(* PLC project GeneratedProgram, SafePLC-Gen SafePLC-Gen Multimodal 1.0 *)
(* stored: creationDateTime 2026-04-25T12:15:41.761626Z *)

PROGRAM GeneratedProgram
  VAR
    TI_2909_Scaled : REAL;
    TT_2909_Scaled : REAL;
    TT_2911_Scaled : REAL;
    TT_2917_Scaled : REAL;
    TI_2917_Scaled : REAL;
    XI_2901A_Scaled : REAL;
    XI_2901B_Scaled : REAL;
    TI_2909_HH_SP : REAL;
    TI_2909_H_SP : REAL;
    TI_2909_L_SP : REAL;
    TI_2909_LL_SP : REAL;
    TI_2909_Deadband : REAL;
    TI_2909_HH : BOOL;
    TI_2909_H : BOOL;
    TI_2909_L : BOOL;
    TI_2909_LL : BOOL;
    TI_2909_HH_Latch : SR;
    TI_2909_LL_Latch : SR;
    TI_2909_HH_Ack : BOOL;
    TI_2909_LL_Ack : BOOL;
    TT_2909_HH_SP : REAL;
    TT_2909_H_SP : REAL;
    TT_2909_L_SP : REAL;
    TT_2909_LL_SP : REAL;
    TT_2909_Deadband : REAL;
    TT_2909_HH : BOOL;
    TT_2909_H : BOOL;
    TT_2909_L : BOOL;
    TT_2909_LL : BOOL;
    TT_2909_HH_Latch : SR;
    TT_2909_LL_Latch : SR;
    TT_2909_HH_Ack : BOOL;
    TT_2909_LL_Ack : BOOL;
    TT_2911_HH_SP : REAL;
    TT_2911_H_SP : REAL;
    TT_2911_L_SP : REAL;
    TT_2911_LL_SP : REAL;
    TT_2911_Deadband : REAL;
    TT_2911_HH : BOOL;
    TT_2911_H : BOOL;
    TT_2911_L : BOOL;
    TT_2911_LL : BOOL;
    TT_2911_HH_Latch : SR;
    TT_2911_LL_Latch : SR;
    TT_2911_HH_Ack : BOOL;
    TT_2911_LL_Ack : BOOL;
    TIC_2911_SP : REAL;
    TIC_2911_Kp : REAL;
    TIC_2911_Ki : REAL;
    TIC_2911_Error : REAL;
    TIC_2911_Integral : REAL;
    TIC_2911_Output : REAL;
    TT_2917_HH_SP : REAL;
    TT_2917_H_SP : REAL;
    TT_2917_L_SP : REAL;
    TT_2917_LL_SP : REAL;
    TT_2917_Deadband : REAL;
    TT_2917_HH : BOOL;
    TT_2917_H : BOOL;
    TT_2917_L : BOOL;
    TT_2917_LL : BOOL;
    TT_2917_HH_Latch : SR;
    TT_2917_LL_Latch : SR;
    TT_2917_HH_Ack : BOOL;
    TT_2917_LL_Ack : BOOL;
    TI_2917_HH_SP : REAL;
    TI_2917_H_SP : REAL;
    TI_2917_L_SP : REAL;
    TI_2917_LL_SP : REAL;
    TI_2917_Deadband : REAL;
    TI_2917_HH : BOOL;
    TI_2917_H : BOOL;
    TI_2917_L : BOOL;
    TI_2917_LL : BOOL;
    TI_2917_HH_Latch : SR;
    TI_2917_LL_Latch : SR;
    TI_2917_HH_Ack : BOOL;
    TI_2917_LL_Ack : BOOL;
    XI_2901A_HH_SP : REAL;
    XI_2901A_H_SP : REAL;
    XI_2901A_L_SP : REAL;
    XI_2901A_LL_SP : REAL;
    XI_2901A_Deadband : REAL;
    XI_2901A_HH : BOOL;
    XI_2901A_H : BOOL;
    XI_2901A_L : BOOL;
    XI_2901A_LL : BOOL;
    XI_2901A_HH_Latch : SR;
    XI_2901A_LL_Latch : SR;
    XI_2901A_HH_Ack : BOOL;
    XI_2901A_LL_Ack : BOOL;
    XI_2901B_HH_SP : REAL;
    XI_2901B_H_SP : REAL;
    XI_2901B_L_SP : REAL;
    XI_2901B_LL_SP : REAL;
    XI_2901B_Deadband : REAL;
    XI_2901B_HH : BOOL;
    XI_2901B_H : BOOL;
    XI_2901B_L : BOOL;
    XI_2901B_LL : BOOL;
    XI_2901B_HH_Latch : SR;
    XI_2901B_LL_Latch : SR;
    XI_2901B_HH_Ack : BOOL;
    XI_2901B_LL_Ack : BOOL;
    LOOP_2917_TRIP : BOOL;
    LOOP_2901A_TRIP : BOOL;
    LOOP_2901B_TRIP : BOOL;
    LOOP_3200_TRIP : BOOL;
    TT_2917_HH_Trip : BOOL;
    TT_2917_LL_Trip : BOOL;
    VSHH_2901A_HH : BOOL;
    VSHH_2901A_LL : BOOL;
    VSHH_2901B_HH : BOOL;
    VSHH_2901B_LL : BOOL;
    ESD_3200_HH : BOOL;
    ESD_3200_LL : BOOL;
    SAFE_STATE : BOOL;
    MotorA_LocalMode : BOOL;
    MotorA_StartCmd : BOOL;
    MotorA_StopCmd : BOOL;
    MotorA_Run : BOOL;
    MotorA_Latch : SR;
    MotorB_LocalMode : BOOL;
    MotorB_StartCmd : BOOL;
    MotorB_StopCmd : BOOL;
    MotorB_Run : BOOL;
    MotorB_Latch : SR;
    StartupDelay : TON;
    System_Alarm : BOOL;
    FirstScan : BOOL;
  END_VAR

            IF FirstScan THEN
    LOOP_2917_TRIP       := TRUE;
    LOOP_2901A_TRIP      := TRUE;
    LOOP_2901B_TRIP      := TRUE;
    LOOP_3200_TRIP       := TRUE;
    SAFE_STATE           := TRUE;
    KV_2904_Out          := 6554;
    MCC_A_Out            := FALSE;
    MCC_B_Out            := FALSE;
    PSD_2917_Out         := FALSE;
    MCC_A_and_MCC_B_Out  := FALSE;
    TIC_2911_Integral    := 0.0;
    FirstScan            := FALSE;
    RETURN;
END_IF;

TI_2909_Scaled  := ((INT_TO_REAL(TI_2909_Raw)  - 6554.0) / (32767.0 - 6554.0)) * 150.0;
TT_2909_Scaled  := ((INT_TO_REAL(TT_2909_Raw)  - 6554.0) / (32767.0 - 6554.0)) * 150.0;
TT_2911_Scaled  := ((INT_TO_REAL(TT_2911_Raw)  - 6554.0) / (32767.0 - 6554.0)) * 150.0;
TT_2917_Scaled  := ((INT_TO_REAL(TT_2917_Raw)  - 6554.0) / (32767.0 - 6554.0)) * 150.0;
TI_2917_Scaled  := ((INT_TO_REAL(TI_2917_Raw)  - 6554.0) / (32767.0 - 6554.0)) * 150.0;
XI_2901A_Scaled := ((INT_TO_REAL(XI_2901A_Raw) - 6554.0) / (32767.0 - 6554.0)) * 100.0;
XI_2901B_Scaled := ((INT_TO_REAL(XI_2901B_Raw) - 6554.0) / (32767.0 - 6554.0)) * 100.0;

TT_2917_HH_Trip := TT_2917_Scaled >= TT_2917_HH_SP;
TT_2917_LL_Trip := TT_2917_Scaled <= TT_2917_LL_SP;
VSHH_2901A_HH   := VSHH_2901A;
VSHH_2901A_LL   := FALSE;
VSHH_2901B_HH   := VSHH_2901B;
VSHH_2901B_LL   := FALSE;
ESD_3200_HH     := ESD_3200;
ESD_3200_LL     := FALSE;

IF TT_2917_HH_Trip OR TT_2917_LL_Trip OR PSD_2917 THEN
    LOOP_2917_TRIP := TRUE;
ELSIF LOOP_2917_TRIP AND MANUAL_RESET
      AND NOT TT_2917_HH_Trip AND NOT TT_2917_LL_Trip AND NOT PSD_2917 THEN
    LOOP_2917_TRIP := FALSE;
END_IF;

IF VSHH_2901A_HH OR VSHH_2901A_LL OR HS_EMERGENCY_STOP_A_2901A THEN
    LOOP_2901A_TRIP := TRUE;
ELSIF LOOP_2901A_TRIP AND MANUAL_RESET
      AND NOT VSHH_2901A_HH AND NOT VSHH_2901A_LL AND NOT HS_EMERGENCY_STOP_A_2901A THEN
    LOOP_2901A_TRIP := FALSE;
END_IF;

IF VSHH_2901B_HH OR VSHH_2901B_LL OR HS_EMERGENCY_STOP_B_2901B THEN
    LOOP_2901B_TRIP := TRUE;
ELSIF LOOP_2901B_TRIP AND MANUAL_RESET
      AND NOT VSHH_2901B_HH AND NOT VSHH_2901B_LL AND NOT HS_EMERGENCY_STOP_B_2901B THEN
    LOOP_2901B_TRIP := FALSE;
END_IF;

IF ESD_3200_HH OR ESD_3200_LL THEN
    LOOP_3200_TRIP := TRUE;
ELSIF LOOP_3200_TRIP AND MANUAL_RESET
      AND NOT ESD_3200_HH AND NOT ESD_3200_LL THEN
    LOOP_3200_TRIP := FALSE;
END_IF;

SAFE_STATE := ESTOP
              OR LOOP_2917_TRIP
              OR LOOP_2901A_TRIP
              OR LOOP_2901B_TRIP
              OR LOOP_3200_TRIP;

IF NOT SAFE_STATE THEN
    TIC_2911_Error    := TIC_2911_SP - TT_2911_Scaled;
    TIC_2911_Integral := TIC_2911_Integral + (TIC_2911_Ki * TIC_2911_Error);
    IF TIC_2911_Integral > 100.0 THEN
        TIC_2911_Integral := 100.0;
    ELSIF TIC_2911_Integral < 0.0 THEN
        TIC_2911_Integral := 0.0;
    END_IF;
    TIC_2911_Output := (TIC_2911_Kp * TIC_2911_Error) + TIC_2911_Integral;
    IF TIC_2911_Output > 100.0 THEN
        TIC_2911_Output := 100.0;
    ELSIF TIC_2911_Output < 0.0 THEN
        TIC_2911_Output := 0.0;
    END_IF;
    KV_2904_Out := REAL_TO_INT(6554.0 + (TIC_2911_Output / 100.0) * (32767.0 - 6554.0));

    MotorA_LocalMode := HS_2901A1;
    IF MotorA_LocalMode THEN
        MotorA_StartCmd := HS_START_STOP_A_2901A;
        MotorA_StopCmd  := NOT HS_START_STOP_A_2901A;
    ELSE
        MotorA_StartCmd := HS_2901A AND HS_2901A2;
        MotorA_StopCmd  := NOT HS_2901A2;
    END_IF;
    MotorA_Latch(S1 := MotorA_StartCmd, R := MotorA_StopCmd);
    MotorA_Run := MotorA_Latch.Q1;

    MotorB_LocalMode := HS_2901B1;
    IF MotorB_LocalMode THEN
        MotorB_StartCmd := HS_START_STOP_B_2901B;
        MotorB_StopCmd  := NOT HS_START_STOP_B_2901B;
    ELSE
        MotorB_StartCmd := HS_2901B AND HS_2901B2;
        MotorB_StopCmd  := NOT HS_2901B2;
    END_IF;
    MotorB_Latch(S1 := MotorB_StartCmd, R := MotorB_StopCmd);
    MotorB_Run := MotorB_Latch.Q1;

    StartupDelay(IN := MotorA_Run OR MotorB_Run, PT := T#3S);

    MCC_A_Out           := MotorA_Run AND StartupDelay.Q;
    MCC_B_Out           := MotorB_Run AND StartupDelay.Q;
    PSD_2917_Out        := TRUE;
    MCC_A_and_MCC_B_Out := MCC_A_Out AND MCC_B_Out;
ELSE
    KV_2904_Out         := 6554;
    MCC_A_Out           := FALSE;
    MCC_B_Out           := FALSE;
    PSD_2917_Out        := FALSE;
    MCC_A_and_MCC_B_Out := FALSE;
    TIC_2911_Integral   := 0.0;
END_IF;

(* TI_2909 four-level alarms *)
IF TI_2909_Scaled >= TI_2909_HH_SP THEN
    TI_2909_HH_Latch.S1 := TRUE;
ELSIF TI_2909_Scaled <= (TI_2909_HH_SP - TI_2909_Deadband) THEN
    TI_2909_HH_Latch.S1 := FALSE;
END_IF;
TI_2909_HH_Latch(S1 := TI_2909_HH_Latch.S1, R := TI_2909_HH_Ack AND (TI_2909_Scaled < TI_2909_HH_SP));
TI_2909_HH := TI_2909_HH_Latch.Q1;
TI_2909_H  := TI_2909_Scaled >= TI_2909_H_SP AND TI_2909_Scaled < TI_2909_HH_SP;
TI_2909_L  := TI_2909_Scaled <= TI_2909_L_SP AND TI_2909_Scaled > TI_2909_LL_SP;
IF TI_2909_Scaled <= TI_2909_LL_SP THEN
    TI_2909_LL_Latch.S1 := TRUE;
ELSIF TI_2909_Scaled >= (TI_2909_LL_SP + TI_2909_Deadband) THEN
    TI_2909_LL_Latch.S1 := FALSE;
END_IF;
TI_2909_LL_Latch(S1 := TI_2909_LL_Latch.S1, R := TI_2909_LL_Ack AND (TI_2909_Scaled > TI_2909_LL_SP));
TI_2909_LL := TI_2909_LL_Latch.Q1;

(* TT_2909 four-level alarms *)
IF TT_2909_Scaled >= TT_2909_HH_SP THEN
    TT_2909_HH_Latch.S1 := TRUE;
ELSIF TT_2909_Scaled <= (TT_2909_HH_SP - TT_2909_Deadband) THEN
    TT_2909_HH_Latch.S1 := FALSE;
END_IF;
TT_2909_HH_Latch(S1 := TT_2909_HH_Latch.S1, R := TT_2909_HH_Ack AND (TT_2909_Scaled < TT_2909_HH_SP));
TT_2909_HH := TT_2909_HH_Latch.Q1;
TT_2909_H  := TT_2909_Scaled >= TT_2909_H_SP AND TT_2909_Scaled < TT_2909_HH_SP;
TT_2909_L  := TT_2909_Scaled <= TT_2909_L_SP AND TT_2909_Scaled > TT_2909_LL_SP;
IF TT_2909_Scaled <= TT_2909_LL_SP THEN
    TT_2909_LL_Latch.S1 := TRUE;
ELSIF TT_2909_Scaled >= (TT_2909_LL_SP + TT_2909_Deadband) THEN
    TT_2909_LL_Latch.S1 := FALSE;
END_IF;
TT_2909_LL_Latch(S1 := TT_2909_LL_Latch.S1, R := TT_2909_LL_Ack AND (TT_2909_Scaled > TT_2909_LL_SP));
TT_2909_LL := TT_2909_LL_Latch.Q1;

(* TT_2911 four-level alarms *)
IF TT_2911_Scaled >= TT_2911_HH_SP THEN
    TT_2911_HH_Latch.S1 := TRUE;
ELSIF TT_2911_Scaled <= (TT_2911_HH_SP - TT_2911_Deadband) THEN
    TT_2911_HH_Latch.S1 := FALSE;
END_IF;
TT_2911_HH_Latch(S1 := TT_2911_HH_Latch.S1, R := TT_2911_HH_Ack AND (TT_2911_Scaled < TT_2911_HH_SP));
TT_2911_HH := TT_2911_HH_Latch.Q1;
TT_2911_H  := TT_2911_Scaled >= TT_2911_H_SP AND TT_2911_Scaled < TT_2911_HH_SP;
TT_2911_L  := TT_2911_Scaled <= TT_2911_L_SP AND TT_2911_Scaled > TT_2911_LL_SP;
IF TT_2911_Scaled <= TT_2911_LL_SP THEN
    TT_2911_LL_Latch.S1 := TRUE;
ELSIF TT_2911_Scaled >= (TT_2911_LL_SP + TT_2911_Deadband) THEN
    TT_2911_LL_Latch.S1 := FALSE;
END_IF;
TT_2911_LL_Latch(S1 := TT_2911_LL_Latch.S1, R := TT_2911_LL_Ack AND (TT_2911_Scaled > TT_2911_LL_SP));
TT_2911_LL := TT_2911_LL_Latch.Q1;

(* TT_2917 four-level alarms *)
IF TT_2917_Scaled >= TT_2917_HH_SP THEN
    TT_2917_HH_Latch.S1 := TRUE;
ELSIF TT_2917_Scaled <= (TT_2917_HH_SP - TT_2917_Deadband) THEN
    TT_2917_HH_Latch.S1 := FALSE;
END_IF;
TT_2917_HH_Latch(S1 := TT_2917_HH_Latch.S1, R := TT_2917_HH_Ack AND (TT_2917_Scaled < TT_2917_HH_SP));
TT_2917_HH := TT_2917_HH_Latch.Q1;
TT_2917_H  := TT_2917_Scaled >= TT_2917_H_SP AND TT_2917_Scaled < TT_2917_HH_SP;
TT_2917_L  := TT_2917_Scaled <= TT_2917_L_SP AND TT_2917_Scaled > TT_2917_LL_SP;
IF TT_2917_Scaled <= TT_2917_LL_SP THEN
    TT_2917_LL_Latch.S1 := TRUE;
ELSIF TT_2917_Scaled >= (TT_2917_LL_SP + TT_2917_Deadband) THEN
    TT_2917_LL_Latch.S1 := FALSE;
END_IF;
TT_2917_LL_Latch(S1 := TT_2917_LL_Latch.S1, R := TT_2917_LL_Ack AND (TT_2917_Scaled > TT_2917_LL_SP));
TT_2917_LL := TT_2917_LL_Latch.Q1;

(* TI_2917 four-level alarms *)
IF TI_2917_Scaled >= TI_2917_HH_SP THEN
    TI_2917_HH_Latch.S1 := TRUE;
ELSIF TI_2917_Scaled <= (TI_2917_HH_SP - TI_2917_Deadband) THEN
    TI_2917_HH_Latch.S1 := FALSE;
END_IF;
TI_2917_HH_Latch(S1 := TI_2917_HH_Latch.S1, R := TI_2917_HH_Ack AND (TI_2917_Scaled < TI_2917_HH_SP));
TI_2917_HH := TI_2917_HH_Latch.Q1;
TI_2917_H  := TI_2917_Scaled >= TI_2917_H_SP AND TI_2917_Scaled < TI_2917_HH_SP;
TI_2917_L  := TI_2917_Scaled <= TI_2917_L_SP AND TI_2917_Scaled > TI_2917_LL_SP;
IF TI_2917_Scaled <= TI_2917_LL_SP THEN
    TI_2917_LL_Latch.S1 := TRUE;
ELSIF TI_2917_Scaled >= (TI_2917_LL_SP + TI_2917_Deadband) THEN
    TI_2917_LL_Latch.S1 := FALSE;
END_IF;
TI_2917_LL_Latch(S1 := TI_2917_LL_Latch.S1, R := TI_2917_LL_Ack AND (TI_2917_Scaled > TI_2917_LL_SP));
TI_2917_LL := TI_2917_LL_Latch.Q1;

(* XI_2901A four-level alarms *)
IF XI_2901A_Scaled >= XI_2901A_HH_SP THEN
    XI_2901A_HH_Latch.S1 := TRUE;
ELSIF XI_2901A_Scaled <= (XI_2901A_HH_SP - XI_2901A_Deadband) THEN
    XI_2901A_HH_Latch.S1 := FALSE;
END_IF;
XI_2901A_HH_Latch(S1 := XI_2901A_HH_Latch.S1, R := XI_2901A_HH_Ack AND (XI_2901A_Scaled < XI_2901A_HH_SP));
XI_2901A_HH := XI_2901A_HH_Latch.Q1;
XI_2901A_H  := XI_2901A_Scaled >= XI_2901A_H_SP AND XI_2901A_Scaled < XI_2901A_HH_SP;
XI_2901A_L  := XI_2901A_Scaled <= XI_2901A_L_SP AND XI_2901A_Scaled > XI_2901A_LL_SP;
IF XI_2901A_Scaled <= XI_2901A_LL_SP THEN
    XI_2901A_LL_Latch.S1 := TRUE;
ELSIF XI_2901A_Scaled >= (XI_2901A_LL_SP + XI_2901A_Deadband) THEN
    XI_2901A_LL_Latch.S1 := FALSE;
END_IF;
XI_2901A_LL_Latch(S1 := XI_2901A_LL_Latch.S1, R := XI_2901A_LL_Ack AND (XI_2901A_Scaled > XI_2901A_LL_SP));
XI_2901A_LL := XI_2901A_LL_Latch.Q1;

(* XI_2901B four-level alarms *)
IF XI_2901B_Scaled >= XI_2901B_HH_SP THEN
    XI_2901B_HH_Latch.S1 := TRUE;
ELSIF XI_2901B_Scaled <= (XI_2901B_HH_SP - XI_2901B_Deadband) THEN
    XI_2901B_HH_Latch.S1 := FALSE;
END_IF;
XI_2901B_HH_Latch(S1 := XI_2901B_HH_Latch.S1, R := XI_2901B_HH_Ack AND (XI_2901B_Scaled < XI_2901B_HH_SP));
XI_2901B_HH := XI_2901B_HH_Latch.Q1;
XI_2901B_H  := XI_2901B_Scaled >= XI_2901B_H_SP AND XI_2901B_Scaled < XI_2901B_HH_SP;
XI_2901B_L  := XI_2901B_Scaled <= XI_2901B_L_SP AND XI_2901B_Scaled > XI_2901B_LL_SP;
IF XI_2901B_Scaled <= XI_2901B_LL_SP THEN
    XI_2901B_LL_Latch.S1 := TRUE;
ELSIF XI_2901B_Scaled >= (XI_2901B_LL_SP + XI_2901B_Deadband) THEN
    XI_2901B_LL_Latch.S1 := FALSE;
END_IF;
XI_2901B_LL_Latch(S1 := XI_2901B_LL_Latch.S1, R := XI_2901B_LL_Ack AND (XI_2901B_Scaled > XI_2901B_LL_SP));
XI_2901B_LL := XI_2901B_LL_Latch.Q1;

System_Alarm :=
    TI_2909_HH_Latch.Q1 OR TI_2909_LL_Latch.Q1 OR TI_2909_H OR TI_2909_L OR
    TT_2909_HH_Latch.Q1 OR TT_2909_LL_Latch.Q1 OR TT_2909_H OR TT_2909_L OR
    TT_2911_HH_Latch.Q1 OR TT_2911_LL_Latch.Q1 OR TT_2911_H OR TT_2911_L OR
    TT_2917_HH_Latch.Q1 OR TT_2917_LL_Latch.Q1 OR TT_2917_H OR TT_2917_L OR
    TI_2917_HH_Latch.Q1 OR TI_2917_LL_Latch.Q1 OR TI_2917_H OR TI_2917_L OR
    XI_2901A_HH_Latch.Q1 OR XI_2901A_LL_Latch.Q1 OR XI_2901A_H OR XI_2901A_L OR
    XI_2901B_HH_Latch.Q1 OR XI_2901B_LL_Latch.Q1 OR XI_2901B_H OR XI_2901B_L OR
    SAFE_STATE;
          
END_PROGRAM

CONFIGURATION Config0
  RESOURCE Res0 ON PLC
    TASK MainTask(INTERVAL := T#20ms, PRIORITY := 0);
    PROGRAM Main : GeneratedProgram;
  END_RESOURCE
END_CONFIGURATION
